// TIA Portal V21 export
// export: Created 2000-01-01T00:00:00.0000000Z, ExportSetting None
TYPE "UDT_HMI_FIO_SortingByHeight"
   STRUCT
      bManualMode { ExternalWritable := 'False'} : Bool;   // TRUE: 手动模式, FALSE: 自动模式
      bStartCmd { ExternalWritable := 'False'} : Bool;   // HMI启动按钮触发
      bStopCmd { ExternalWritable := 'False'} : Bool;   // HMI停止按钮触发
      bResetCmd { ExternalWritable := 'False'} : Bool;   // HMI故障复位触发
      bManualEntryConv { ExternalWritable := 'False'} : Bool;   // 手动驱动入口传送带
      bManualExitConv { ExternalWritable := 'False'} : Bool;   // 手动驱动出口传送带
      bManualPusherHigh { ExternalWritable := 'False'} : Bool;   // 手动伸出高件推杆
      bManualPusherLow { ExternalWritable := 'False'} : Bool;   // 手动伸出低件推杆
      tTransferTimeout { ExternalWritable := 'False'} : Time;   // 分拣滑道传送超时时间（默认 T#8s）
      tPusherHoldTime { ExternalWritable := 'False'} : Time;   // 推杆推出保持时间（默认 T#800ms）
      iCurrentStep { ExternalWritable := 'False'} : Int;   // 状态反馈：当前顺控步号
      diHighSortedCount { ExternalWritable := 'False'} : DInt;   // 状态反馈：已分拣高件计数
      diLowSortedCount { ExternalWritable := 'False'} : DInt;   // 状态反馈：已分拣低件计数
      bRunning { ExternalWritable := 'False'} : Bool;   // 状态反馈：系统运行中
      bFault { ExternalWritable := 'False'} : Bool;   // 状态反馈：分拣超时或急停故障
      wStatus { ExternalWritable := 'False'} : Word;   // 状态码：16#0000运行正常, 16#7000待机, 16#8401分拣传送超时, 16#8402急停触发
   END_STRUCT;
END_TYPE
